(* IEC 61131-3 sources: Jacob-Formschaumtechnik-ISEL-CNC-Retrofit/twincat/PLC/src/3_Cnc, 2 files *)

(* ---- FB_CncMirror.st ---- *)
(* CNC-Spiegel fuer die HMI (GVL_HmiCnc). Solange TF5200/TF5310 fehlen, arbeitet er als Simulation:
   Overrides werden begrenzt, Programm laden und Tabellen schreiben nur im Stillstand,
   sonst bTableWriteRejected. Spaeter speist die CNC (Tc2_CncHli) dieselben Felder. Positionen bleiben
   in der Simulation stehen (keine Bewegung). Befund 23. *)
FUNCTION_BLOCK FB_CncMirror
VAR_INPUT
    bStandstill : BOOL;      (* kein Programm aktiv, kein Halt *)
END_VAR
VAR_IN_OUT
    stCmd : ST_HmiCncCmd;
    stSts : ST_HmiCncSts;
END_VAR
VAR
    rtLoad  : R_TRIG;
    rtWrite : R_TRIG;
    rtWcs   : R_TRIG;
    nIdx    : INT;
    nLimit  : UINT := 25;      (* wirksame Inbetriebnahme-Begrenzung in %, nach dem Anlauf immer 25 *)
    rtWcsWrite : R_TRIG;
END_VAR

rtLoad(CLK := stCmd.bProgramLoad);
rtWrite(CLK := stCmd.bTableWrite);
rtWcs(CLK := stCmd.bWcsSetCurrent);

(* Overrides begrenzen, die SPS entscheidet *)
(* Inbetriebnahme-Begrenzung: Absenken sofort, Anheben nur im Stillstand, immer 1..100 % *)
IF stCmd.nSpeedLimitPct < 1 THEN
    nLimit := 1;
ELSIF stCmd.nSpeedLimitPct < nLimit THEN
    nLimit := MIN(stCmd.nSpeedLimitPct, 100);
ELSIF stCmd.nSpeedLimitPct > nLimit AND bStandstill THEN
    nLimit := MIN(stCmd.nSpeedLimitPct, 100);
END_IF
stSts.nSpeedLimitActivePct := nLimit;

stSts.nOvrFeed    := MIN(stCmd.nOvrFeed, 120) * nLimit / 100;
stSts.nOvrRapid   := MIN(stCmd.nOvrRapid, 100) * nLimit / 100;
stSts.nOvrSpindle := LIMIT(50, stCmd.nOvrSpindle, 120);

rtWcsWrite(CLK := stCmd.bWcsTableWrite);
IF rtLoad.Q OR rtWrite.Q OR rtWcs.Q OR rtWcsWrite.Q THEN
    stSts.bTableWriteOk := FALSE;
    stSts.bTableWriteRejected := FALSE;
END_IF

IF rtLoad.Q THEN
    IF bStandstill THEN
        stSts.sProgramName := stCmd.sProgramSelect;
        stSts.bProgramLoaded := stCmd.sProgramSelect <> '';
        stSts.bTableWriteOk := TRUE;
    ELSE
        stSts.bTableWriteRejected := TRUE;
    END_IF
END_IF

(* G-16: Werkzeugtabelle und Nullpunkte haben getrennte Schreibimpulse, damit das Speichern der Werkzeuge
   nie die Nullpunkte ueberschreibt *)
IF rtWrite.Q THEN
    IF bStandstill THEN
        stSts.aTool := stCmd.aTool;
        stSts.bTableWriteOk := TRUE;
    ELSE
        stSts.bTableWriteRejected := TRUE;
    END_IF
END_IF

IF rtWcsWrite.Q THEN
    IF bStandstill THEN
        stSts.aWcs := stCmd.aWcs;
        stSts.bTableWriteOk := TRUE;
    ELSE
        stSts.bTableWriteRejected := TRUE;
    END_IF
END_IF

IF rtWcs.Q THEN
    nIdx := UINT_TO_INT(stSts.nActWcs);
    IF bStandstill AND nIdx >= 54 AND nIdx <= 59 THEN
        stSts.aWcs[nIdx].rX := stSts.aAxis[1].rActPosMach;
        stSts.aWcs[nIdx].rY := stSts.aAxis[2].rActPosMach;
        stSts.aWcs[nIdx].rZ := stSts.aAxis[3].rActPosMach;
        stCmd.aWcs[nIdx] := stSts.aWcs[nIdx];
        stSts.bTableWriteOk := TRUE;
    ELSE
        stSts.bTableWriteRejected := TRUE;
    END_IF
END_IF
END_FUNCTION_BLOCK

(* ---- FB_MFunctions.st ---- *)
(* Hilfsfunktionen aus dem NC-Programm (M-Codes). Die Zuordnung orientiert sich an der
   isel-G-/M-Code-Liste (Klaerungsliste Funktionen 2.7). Welche M-Codes der Kunde tatsaechlich
   braucht, bestimmt das Lastenheft (2.8.2). Die Anbindung an die CNC (Tc2_CncHli) folgt.
   Gutachten G-03: M3/M4 wird erst quittiert, wenn die Spindel laeuft (oder bewusst gesperrt ist: Einrichten,
   Trockenlauf). Ein M-Code ohne Ausfuehrungsmoeglichkeit und ein unbekannter M-Code werden nicht quittiert.
   G-04: Das Vakuum bleibt bei Abbruch und NOT-HALT gehalten (Werkstueckspannung), es geht mit M11, M30/M2 oder von Hand aus. *)
FUNCTION_BLOCK FB_MFunctions
VAR_INPUT
    nMCode      : INT;          (* aktive M-Funktion aus der CNC, 0 = keine *)
    bMStrobe    : BOOL;         (* CNC wartet auf Quittung *)
    bSpindleOk  : BOOL;
    bAuxOk      : BOOL;
    bReset      : BOOL;         (* Abbruch, R3/R4, NOT-HALT, Programmende: gehaltene M-Zustaende loeschen (ausser Vakuum) *)
    bOptStop    : BOOL;         (* optionaler Halt M1 aktiv (aus der HMI) *)
    bSpindleRunning : BOOL;     (* Spindel hat Drehzahl erreicht *)
    bSpindleSkip    : BOOL;     (* Einrichten/Trockenlauf: Spindel bewusst aus, M3/M4 ohne Start quittieren *)
END_VAR
VAR_OUTPUT
    bSpindleCw    : BOOL;       (* M3 *)
    bSpindleCcw   : BOOL;       (* M4 *)
    bExtraction   : BOOL;       (* M43 ein, M44 aus [Annahme: Belegung klaeren] *)
    bBlowAir      : BOOL;       (* M8 ein, M9 aus *)
    bVacuum       : BOOL;       (* M10 ein, M11 aus *)
    bToolChangeReq: BOOL;       (* M6: manuelle Aufforderung am Panel *)
    bProgramHalt  : BOOL;       (* M0 *)
    bAck          : BOOL;       (* Quittung an die CNC *)
    bUnknown      : BOOL;       (* unbekannter M-Code: nicht quittiert *)
END_VAR
VAR
    rtStrobe    : R_TRIG;
    bWaitSpindle: BOOL;         (* Quittung zurueckgehalten, bis die Spindel laeuft *)
    bBlockAck   : BOOL;         (* M-Code nicht ausfuehrbar: nie quittieren *)
END_VAR

rtStrobe(CLK := bMStrobe);
bUnknown := FALSE; bToolChangeReq := FALSE; bProgramHalt := FALSE;

IF bReset THEN
    bSpindleCw := FALSE; bSpindleCcw := FALSE; bExtraction := FALSE; bBlowAir := FALSE;
    bWaitSpindle := FALSE;      (* G-04: bVacuum bleibt gehalten *)
END_IF
IF NOT bMStrobe THEN
    bWaitSpindle := FALSE; bBlockAck := FALSE;
END_IF

IF rtStrobe.Q AND NOT bReset THEN
    CASE nMCode OF
        0:  bProgramHalt := TRUE;
        1:  IF bOptStop THEN bProgramHalt := TRUE; END_IF
        3:  IF bSpindleSkip THEN
                bSpindleCw := FALSE; bSpindleCcw := FALSE;     (* Spindel bewusst aus, Programm laeuft weiter *)
            ELSIF bSpindleOk THEN
                bSpindleCw := TRUE; bSpindleCcw := FALSE; bWaitSpindle := TRUE;
            ELSE
                bBlockAck := TRUE;                                (* nicht ausfuehrbar: nicht quittieren *)
            END_IF
        4:  IF bSpindleSkip THEN
                bSpindleCw := FALSE; bSpindleCcw := FALSE;
            ELSIF bSpindleOk THEN
                bSpindleCcw := TRUE; bSpindleCw := FALSE; bWaitSpindle := TRUE;
            ELSE
                bBlockAck := TRUE;
            END_IF
        5:  bSpindleCw := FALSE; bSpindleCcw := FALSE;
        6:  bToolChangeReq := TRUE;
        8:  IF bAuxOk THEN bBlowAir := TRUE; END_IF
        9:  bBlowAir := FALSE;
        10: IF bAuxOk THEN bVacuum := TRUE; END_IF
        11: bVacuum := FALSE;
        2, 30: bSpindleCw := FALSE; bSpindleCcw := FALSE; bBlowAir := FALSE; bExtraction := FALSE; bVacuum := FALSE;
        43: IF bAuxOk THEN bExtraction := TRUE; END_IF
        44: bExtraction := FALSE;
    ELSE
        bUnknown := TRUE; bBlockAck := TRUE;
    END_CASE
END_IF

IF bWaitSpindle AND (bSpindleRunning OR bSpindleSkip) THEN bWaitSpindle := FALSE; END_IF

(* Quittung bleibt stehen, bis die CNC den Strobe zurueckgenommen hat; zurueckgehalten bei M3/M4 bis die Spindel laeuft *)
bAck := bMStrobe AND NOT bWaitSpindle AND NOT bBlockAck;
END_FUNCTION_BLOCK
